(* IEC 61131-3 sources: kns-port-domestic/tools/plcopen/tests/fixtures/constructs/src/POUs/Devices/FB_DeviceBase, 4 files *)

(* ---- FB_DeviceBase.decl.st ---- *)
// Назначение: абстрактная база устройств — режим, отказ, квитирование
// Автор:      <ИМЯ ФАМИЛИЯ>
// Версия:     0.1.0
// Документ:   docs/plcopen.md
{attribute 'reflection'}
FUNCTION_BLOCK ABSTRACT FB_DeviceBase IMPLEMENTS I_Device
VAR_INPUT
    xReset : BOOL;
END_VAR
VAR_OUTPUT
    xFault : BOOL;
END_VAR
VAR
    eModeInt : E_Mode := E_Mode.OutOfService;
    {attribute 'hide'}
    xFaultInt : BOOL;
END_VAR
VAR_STAT
    uiInstances : UINT;
END_VAR

(* ---- FB_DeviceBase.impl.st ---- *)
// общая логика базы: сброс по входу
IF xReset THEN
    Reset(xForce := FALSE);
END_IF
xFault := xFaultInt;

(* ---- Reset.method.decl.st ---- *)
// Сброс отказа
METHOD PUBLIC Reset : BOOL
VAR_INPUT
    xForce : BOOL;
END_VAR

(* ---- SetFault.method.decl.st ---- *)
// Установить отказ (только для наследников)
METHOD PROTECTED SetFault
VAR_INPUT
    xValue : BOOL;
END_VAR
